FUNCTION_BLOCK Heater
VAR_INPUT
	iWaterTemp : REAL;
END_VAR
VAR_OUTPUT
	oHeaterEnable : BOOL;
	oHeaterPower : REAL;
END_VAR
VAR_IN_OUT
	ioHeatStruct : THeater;
END_VAR
VAR
	pidParameters : ST_CTRL_PID_PARAMS;
	pidMode : E_CTRL_MODE;      // ACTIVE when heater is enabled, RESET otherwise
END_VAR

pidParameters.fKp := 1.196; //P
pidParameters.tTn := T#75.798S; //I
pidParameters.tTv := T#0S; //D
pidParameters.tCtrlCycleTime := T#200MS;
pidParameters.tTaskCycleTime := T#100MS;
pidParameters.fOutMaxLimit := 100;
pidParameters.fOutMinLimit := 0;
pidParameters.bDInTheFeedbackPath := FALSE;
pidParameters.bPInTheFeedbackPath := FALSE;
pidParameters.bARWOnIPartOnly := FALSE;
pidParameters.tTd := T#100MS; 


// PID runs only when heater is enabled - otherwise it is held in reset,
// so the integral part doesn't wind up while heating is off (no overshoot after start)
IF ioHeatStruct.State.EnableOut THEN
	pidMode := E_CTRL_MODE.eCTRL_MODE_ACTIVE;
ELSE
	pidMode := E_CTRL_MODE.eCTRL_MODE_RESET;
END_IF;

ioHeatStruct.PID(
	fSetpointValue := ioHeatStruct.ParamHeatingSetPointAutomat, 
	fActualValue := iWaterTemp, 
	fManSyncValue := ioHeatStruct.ParamHeatingPowerManual,
	bSync := ioHeatStruct.State.ManCtrl,
	eMode := pidMode, // automatic mode of PID component
	stParams := pidParameters);

ioHeatStruct.State.HeatingOut := ioHeatStruct.PID.fOut;

	 
{region "Manual/Automat"}
// switching state of engine - automatic or manual control (default state is manual)
	IF ioHeatStruct.Cmd.ManCtrl THEN
      	ioHeatStruct.State.ManCtrl := TRUE;
		ioHeatStruct.State.AutCtrl := FALSE;
	ELSIF ioHeatStruct.Cmd.AutCtrl THEN
        ioHeatStruct.State.ManCtrl := FALSE;
		ioHeatStruct.State.AutCtrl := TRUE; 
    END_IF;
		 
	IF (NOT ioHeatStruct.State.AutCtrl AND NOT ioHeatStruct.State.ManCtrl) THEN
		ioHeatStruct.State.ManCtrl := TRUE;
	END_IF

	ioHeatStruct.Cmd.ManCtrl := FALSE;
	ioHeatStruct.Cmd.AutCtrl := FALSE;
{endregion}
	 
 
{region "ManCtrl"}
	// processing manual actions - if command is processed, it is set to FALSE even if can't be processed
	// Heater commands are turn off (stop) and turn on (start) and power level
	IF ioHeatStruct.State.ManCtrl THEN
		IF ioHeatStruct.Cmd.TurnOnMan AND NOT ioHeatStruct.State.GenErr THEN
			ioHeatStruct.State.EnableOut := TRUE;
		ELSIF ioHeatStruct.Cmd.TurnOffMan THEN
			ioHeatStruct.State.EnableOut := FALSE;
		END_IF
    END_IF;
	ioHeatStruct.Cmd.TurnOnMan := FALSE;
	ioHeatStruct.Cmd.TurnOffMan := FALSE;
{endregion}
 
{region "AutCtrl"}
	//if request to run in automatic mode set outputs to right states if MAR
	//AutoRequest shouldn't be reseted to false state
    IF ioHeatStruct.State.AutCtrl THEN
		IF ioHeatStruct.Cmd.Req2RunAutCtrl AND NOT ioHeatStruct.State.GenErr THEN
			ioHeatStruct.State.EnableOut := TRUE;
		ELSIF NOT ioHeatStruct.Cmd.Req2RunAutCtrl THEN
			ioHeatStruct.State.EnableOut := FALSE;
		END_IF
    END_IF;
{endregion}
 
{region "Error states"}
	// if water temperature is too high, stop heating and generate error
	IF iWaterTemp > 90 THEN
		ioHeatStruct.State.EnableOut := FALSE;
		ioHeatStruct.State.GenErr := TRUE;
	ELSIF iWaterTemp < 85 THEN
		ioHeatStruct.State.GenErr := FALSE;
	END_IF
	ioHeatStruct.State.Err := ioHeatStruct.State.GenErr;
{endregion}
	 
 IF NOT ioHeatStruct.State.EnableOut THEN
    ioHeatStruct.State.HeatingOut := 0;
ELSIF ioHeatStruct.State.ManCtrl THEN
    ioHeatStruct.State.HeatingOut := ioHeatStruct.ParamHeatingPowerManual;
ELSE
    ioHeatStruct.State.HeatingOut := ioHeatStruct.PID.fOut;
END_IF;
 
oHeaterPower := ioHeatStruct.State.HeatingOut;
oHeaterEnable := ioHeatStruct.State.EnableOut;

END_FUNCTION_BLOCK

(* stored: Version 1.1.0.1, ProductVersion 3.1.4026.21
   POU Heater: Id {fe81cd62-8fb3-4eb5-8579-8abf8e5327d3}, SpecialFunc None *)
